{attribute 'qualified_only'}
{attribute 'strict'}
TYPE E_CIP_Type :
(
	NotSelected := 0,
	R_Water,
	Detergent,
	Full
);
END_TYPE

(* stored: Version 1.1.0.1, ProductVersion 3.1.4024.12
   DUT E_CIP_Type: Id {8bb3870c-9424-4138-a985-6a3d7c6b591f} *)
